{attribute 'pack_mode' := '1'}
TYPE ST_Sample :
STRUCT
    nId : UDINT;
    sName : STRING(31);
END_STRUCT
END_TYPE

(* stored: Version 1.1.0.1, ProductVersion 3.1.4024.12
   DUT ST_Sample: Id {11111111-2222-3333-4444-666666666666} *)
